// TIA Portal V21 export
// export: Created 2026-11-08T19:42:31.1843385Z, ExportSetting WithDefaults, DisplayName Totally Integrated Automation Portal, DisplayVersion V21 Update 3, DisplayName STEP 7 Professional, DisplayVersion V21 Update 3, DisplayName STEP 7 Safety, DisplayVersion V21, DisplayName Tech WebApplication, DisplayVersion V21, DisplayName WinCC Basic/Comfort/Advanced, DisplayVersion V21 Update 3, DisplayName WinCC Unified, DisplayVersion V21 Update 3
VAR_GLOBAL   // PLC tag table "TagTable_1"
   Tag_Bool_1 AT %M0.0 : Bool;   // Test
END_VAR
